Fanuc KAREL source: compact_preamble.KL

PROGRAM KX00033
%UNINITVARS
%NOLOCKGROUP
VAR
I:INTEGER;J:INTEGER;B:BOOLEAN
F : FILE
S : STRING[80]
P : XYZWPR
BEGIN
I=1
END KX00033
